Fanuc KAREL source: KX00005.KL

PROGRAM KX00005
%NOLOCKGROUP
VAR
  I: INTEGER
  J: INTEGER
  B: BOOLEAN
  F: FILE
  S: STRING[80]
  P: XYZWPR
BEGIN
  OPEN FILE F ('RW', 'MD:KFSAMPLE.DT')
  CANCEL FILE F
  CLOSE FILE F
END KX00005
